TYPE "ST_PersistResult"
VERSION : 0.1
   STRUCT
      Ok : Bool;
      Found : Bool;
      Lost : Bool;
      Length : UDInt;
      ErrorId : UDInt;
   END_STRUCT;

END_TYPE

